INTERFACE I_SafetyController

PROPERTY EStopOK : BOOL
GET
END_GET
END_PROPERTY

END_INTERFACE

(* stored: Version 1.1.0.1
   Itf I_SafetyController: Id {75cc1dc0-1fe0-0a83-16f9-f86bc902e86f}
   Property EStopOK: Id {2f4df65d-4a99-0047-0aa9-2b7b567f1a9c}
   Get Get: Id {f3af02b7-4557-0a7f-3fff-5ff38992b042} *)
